(* PLC project g_traffic_light_clean, Anonymous Benchmark Suite 1.0 *)
(* stored: creationDateTime 2026-07-09T00:00:00 *)

PROGRAM g_traffic_light_clean
  VAR_INPUT
    ns_req : BOOL;
    ew_req : BOOL;
    maint : BOOL;
  END_VAR
  VAR_OUTPUT
    ns_green : BOOL;
    ew_green : BOOL;
  END_VAR

(* LD diagram, written out as Structured Text *)
ns_green := NOT ew_req AND ns_req;
ew_green := ew_req;
END_PROGRAM

CONFIGURATION Config0
  RESOURCE Res0 ON PLC
    TASK tcyclic(INTERVAL := T#10ms, PRIORITY := 0);
    PROGRAM inst0 WITH tcyclic : g_traffic_light_clean;
  END_RESOURCE
END_CONFIGURATION
